Omron CX-Programmer project NewProject (CX-Programmer 9.73)

# PLC NewPLC1: CP1E NA

## Global symbols (name address type ; comment)
PB_START 0.00 BOOL  ; Push Button Start Sistem
PB_STOP 0.01 BOOL  ; Push Button Stop Sistem
SYS_RUN W0.00 BOOL  ; Status Sistem Aktif
LAMPU_MERAH 100.00 BOOL  ; Output Lampu Merah
LAMPU_KUNING 100.01 BOOL  ; Output Lampu Kuning
LAMPU_HIJAU 100.02 BOOL  ; Output Lampu Hijau
T_MERAH_TOTAL T000 BOOL  ; Timer Merah Total (3.0s)
T_MERAH_PRE_KUNING T001 BOOL  ; Timer Merah sisa 1s (2.0s)
T_HIJAU_TOTAL T002 BOOL  ; Timer Hijau Total (3.0s)
T_HIJAU_PRE_KUNING T003 BOOL  ; Timer Hijau sisa 1s (2.0s)

## Program NewProgram1 (cyclic task 0)

### Section TrafficLight

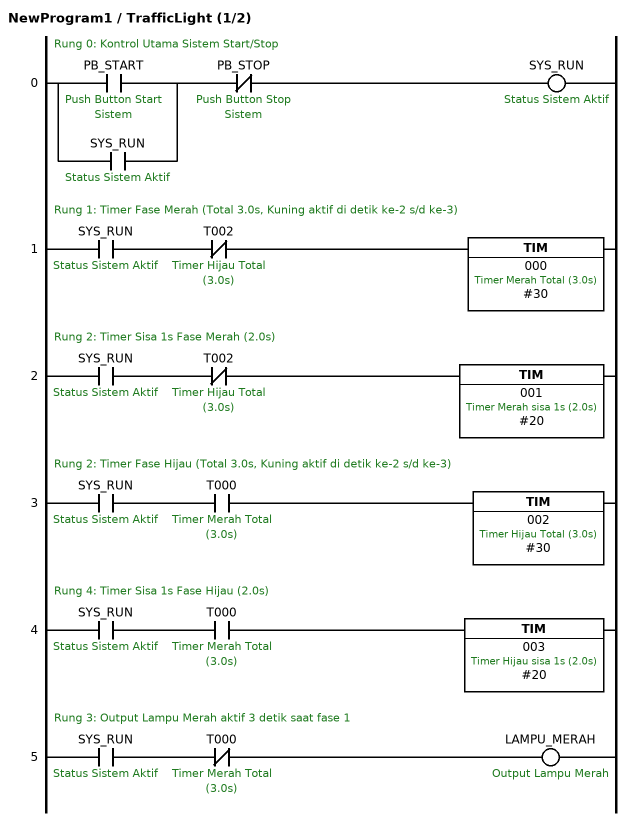
; rung 0: Rung 0: Kontrol Utama Sistem Start/Stop
LD PB_START  ; Push Button Start Sistem
OR SYS_RUN  ; Status Sistem Aktif
ANDNOT PB_STOP  ; Push Button Stop Sistem
OUT SYS_RUN  ; Status Sistem Aktif
; rung 1: Rung 1: Timer Fase Merah (Total 3.0s, Kuning aktif di detik ke-2 s/d ke-3)
LD SYS_RUN  ; Status Sistem Aktif
ANDNOT T002  ; Timer Hijau Total (3.0s)
TIM 000 #30  ; Timer Merah Total (3.0s)
; rung 2: Rung 2: Timer Sisa 1s Fase Merah (2.0s)
LD SYS_RUN  ; Status Sistem Aktif
ANDNOT T002  ; Timer Hijau Total (3.0s)
TIM 001 #20  ; Timer Merah sisa 1s (2.0s)
; rung 3: Rung 2: Timer Fase Hijau (Total 3.0s, Kuning aktif di detik ke-2 s/d ke-3)
LD SYS_RUN  ; Status Sistem Aktif
AND T000  ; Timer Merah Total (3.0s)
TIM 002 #30  ; Timer Hijau Total (3.0s)
; rung 4: Rung 4: Timer Sisa 1s Fase Hijau (2.0s)
LD SYS_RUN  ; Status Sistem Aktif
AND T000  ; Timer Merah Total (3.0s)
TIM 003 #20  ; Timer Hijau sisa 1s (2.0s)
; rung 5: Rung 3: Output Lampu Merah aktif 3 detik saat fase 1
LD SYS_RUN  ; Status Sistem Aktif
ANDNOT T000  ; Timer Merah Total (3.0s)
OUT LAMPU_MERAH  ; Output Lampu Merah

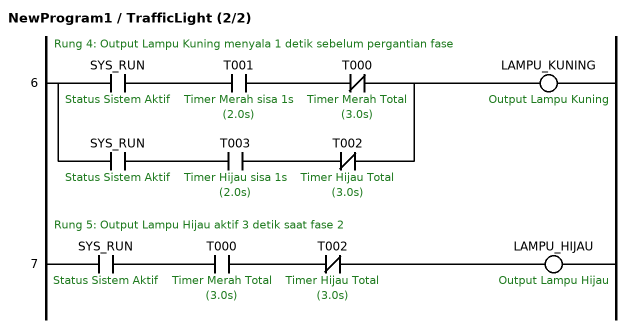
; rung 6: Rung 4: Output Lampu Kuning menyala 1 detik sebelum pergantian fase
LD SYS_RUN  ; Status Sistem Aktif
AND T001  ; Timer Merah sisa 1s (2.0s)
ANDNOT T000  ; Timer Merah Total (3.0s)
LD SYS_RUN  ; Status Sistem Aktif
AND T003  ; Timer Hijau sisa 1s (2.0s)
ANDNOT T002  ; Timer Hijau Total (3.0s)
ORLD
OUT LAMPU_KUNING  ; Output Lampu Kuning
; rung 7: Rung 5: Output Lampu Hijau aktif 3 detik saat fase 2
LD SYS_RUN  ; Status Sistem Aktif
AND T000  ; Timer Merah Total (3.0s)
ANDNOT T002  ; Timer Hijau Total (3.0s)
OUT LAMPU_HIJAU  ; Output Lampu Hijau

### Section END
; rung 0
END(001)